FUNCTION F_DECODE_COMMAND : T_COMMAND
VAR_INPUT
	eCommand: E_COMMAND;
	sCommandData:STRING(255);
END_VAR
VAR

END_VAR

CASE eCommand OF
	E_COMMAND.RALARM:
		F_DECODE_COMMAND.NAME:='RALARM';
		F_DECODE_COMMAND.nData:=0;
	E_COMMAND.RPOSJ:
		F_DECODE_COMMAND.NAME:='RPOSJ';
		F_DECODE_COMMAND.nData:=0;
	E_COMMAND.RPOSC:
		F_DECODE_COMMAND.NAME:='RPOSC';
		F_DECODE_COMMAND.nData:=2;
	E_COMMAND.RSTATS:
		F_DECODE_COMMAND.NAME:='RSTATS';
		F_DECODE_COMMAND.nData:=0;

	E_COMMAND.RJSEQ:
		F_DECODE_COMMAND.NAME:='RJSEQ';
		F_DECODE_COMMAND.nData:=0;
	E_COMMAND.JWAIT:(*NOT SUPPORTED*)
		F_DECODE_COMMAND.NAME:='JWAIT';
		F_DECODE_COMMAND.nData:=1;
	E_COMMAND.RGROUP:
		F_DECODE_COMMAND.NAME:='RGROUP';
		F_DECODE_COMMAND.nData:=0;
	E_COMMAND.RJDIR:
		F_DECODE_COMMAND.NAME:='RJDIR';
		F_DECODE_COMMAND.nData:=1;
	E_COMMAND.RUFRAME:
		F_DECODE_COMMAND.NAME:='RUFRAME';
		F_DECODE_COMMAND.nData:=1;
	E_COMMAND.SAVEV:
		F_DECODE_COMMAND.NAME:='SAVEV';
		F_DECODE_COMMAND.nData:=2;
	E_COMMAND.HOLD:
		F_DECODE_COMMAND.NAME:='HOLD';
		F_DECODE_COMMAND.nData:=1;
	E_COMMAND.RESET:
		F_DECODE_COMMAND.NAME:='RESET';
		F_DECODE_COMMAND.nData:=0;
	E_COMMAND.CANCEL:
		F_DECODE_COMMAND.NAME:='CANCEL';
		F_DECODE_COMMAND.nData:=0;
	E_COMMAND.MODE:
		F_DECODE_COMMAND.NAME:='MODE';
		F_DECODE_COMMAND.nData:=1;
	E_COMMAND.CYCLE:
		F_DECODE_COMMAND.NAME:='CYCLE';
		F_DECODE_COMMAND.nData:=1;
	E_COMMAND.SVON:
		F_DECODE_COMMAND.NAME:='SVON';
		F_DECODE_COMMAND.nData:=1;
	E_COMMAND.HLOCK:
		F_DECODE_COMMAND.NAME:='HLOCK';
		F_DECODE_COMMAND.nData:=1;
	E_COMMAND.MDSP:
		F_DECODE_COMMAND.NAME:='MDSP';
		F_DECODE_COMMAND.nData:=1;
	E_COMMAND.CGROUP:
		F_DECODE_COMMAND.NAME:='CGROUP';
		F_DECODE_COMMAND.nData:=2;
	E_COMMAND.CTASK:
		F_DECODE_COMMAND.NAME:='CTASK';
		F_DECODE_COMMAND.nData:=1;
	E_COMMAND.START:
		F_DECODE_COMMAND.NAME:='START';
		F_DECODE_COMMAND.nData:=0;
	E_COMMAND.START2:
		F_DECODE_COMMAND.NAME:='START';
		F_DECODE_COMMAND.nData:=1;
	E_COMMAND.MOVJ:
		F_DECODE_COMMAND.NAME:='MOVJ';
		F_DECODE_COMMAND.nData:=16;
	E_COMMAND.MOVL:
		F_DECODE_COMMAND.NAME:='MOVL';
		F_DECODE_COMMAND.nData:=17;
	E_COMMAND.IMOV:
		F_DECODE_COMMAND.NAME:='IMOV';
		F_DECODE_COMMAND.nData:=17;
	E_COMMAND.PMOVJ:
		F_DECODE_COMMAND.NAME:='PMOVJ';
		F_DECODE_COMMAND.nData:=14;
	E_COMMAND.PMOVL:
		F_DECODE_COMMAND.NAME:='PMOVL';
		F_DECODE_COMMAND.nData:=15;
	E_COMMAND.DELETE:
		F_DECODE_COMMAND.NAME:='DELETE';
		F_DECODE_COMMAND.nData:=1;
	E_COMMAND.CVTRJ:
		F_DECODE_COMMAND.NAME:='CVTRJ';
		F_DECODE_COMMAND.nData:=2;
	E_COMMAND.CVTSJ:
		F_DECODE_COMMAND.NAME:='CVTSJ';
		F_DECODE_COMMAND.nData:=3;
	E_COMMAND.WUFRAME:
		F_DECODE_COMMAND.NAME:='WUFRAME';
		F_DECODE_COMMAND.nData:=29;
	E_COMMAND.LOADV:
		F_DECODE_COMMAND.NAME:='LOADV';
		F_DECODE_COMMAND.nData:=3;
	E_COMMAND.LOADV2:
		F_DECODE_COMMAND.NAME:='LOADV';
		F_DECODE_COMMAND.nData:=12;
	E_COMMAND.SETMJ:
		F_DECODE_COMMAND.NAME:='SETMJ';
		F_DECODE_COMMAND.nData:=1;
	E_COMMAND.JSEQ:
		F_DECODE_COMMAND.NAME:='JSEQ';
		F_DECODE_COMMAND.nData:=2;
	E_COMMAND.IOREAD:
		F_DECODE_COMMAND.NAME:='IOREAD';
		F_DECODE_COMMAND.nData:=2;
	E_COMMAND.IOWRITE:
		F_DECODE_COMMAND.NAME:='IOWRITE';
		F_DECODE_COMMAND.nData:=1;
	E_COMMAND.IOWRITE2:
		F_DECODE_COMMAND.NAME:='IOWRITE';
		F_DECODE_COMMAND.nData:=2;
	E_COMMAND.IOWRITE3:
		F_DECODE_COMMAND.NAME:='IOWRITE';
		F_DECODE_COMMAND.nData:=3;
	E_COMMAND.IOWRITE4:
		F_DECODE_COMMAND.NAME:='IOWRITE';
		F_DECODE_COMMAND.nData:=4;
	E_COMMAND.IOWRITE5:
		F_DECODE_COMMAND.NAME:='IOWRITE';
		F_DECODE_COMMAND.nData:=5;
	E_COMMAND.IOWRITE6:
		F_DECODE_COMMAND.NAME:='IOWRITE';
		F_DECODE_COMMAND.nData:=6;
	E_COMMAND.IOWRITE7:
		F_DECODE_COMMAND.NAME:='IOWRITE';
		F_DECODE_COMMAND.nData:=7;
	E_COMMAND.IOWRITE8:
		F_DECODE_COMMAND.NAME:='IOWRITE';
		F_DECODE_COMMAND.nData:=8;
	E_COMMAND.IOWRITE9:
		F_DECODE_COMMAND.NAME:='IOWRITE';
		F_DECODE_COMMAND.nData:=9;
	E_COMMAND.IOWRITE10:
		F_DECODE_COMMAND.NAME:='IOWRITE';
		F_DECODE_COMMAND.nData:=10;
END_CASE;

IF	F_DECODE_COMMAND.nData>0	THEN
	F_DECODE_COMMAND.SIZE:=FIND(sCommandData,'$R');
ELSE
	F_DECODE_COMMAND.SIZE:=0;
END_IF;

END_FUNCTION

(* stored: Version 1.1.0.1, ProductVersion 3.1.4024.16
   POU F_DECODE_COMMAND: Id {0e65f4ec-f4c0-4339-8fe3-300583162c1e}, SpecialFunc None *)
